DATA_BLOCK "Tgp_GlobalTemplateFB_LAD"
{ S7_Optimized_Access := 'TRUE' }
VERSION : 0.1
"Tgp_TemplateFB_LAD"
BEGIN
END_DATA_BLOCK
